// TIA Portal V19 export
VAR_GLOBAL   // PLC tag table "Default tag table"
   Simular AT %M100.1 : Bool;
   Test AT %M100.2 : Bool;
   OpContinue AT %M100.0 : Bool;
   EM_Start AT %M0.0 : Bool;
   Tag_1 AT %MW200 : Word;
END_VAR
